FUNCTION_BLOCK basicInversorATV600 (* Inversor ATV600 por Modbus TCP generico: registradores brutos para grandezas e palavras de escrita *)
  (* Standard: 61499-2 *)
  (* Version 1.1, 27/10/2026, Hidryco, Hidryco, 1.1: VELOCIDADE_PCT (leitura) entre LSP 3105 = 0 %% e HSP 3104 = 100 %%. 1.0: Motor_Generico com ATV600 por MODBUSGENTCPS (unit 248): RFR, LCR, UOP, OPR, OTR, LFT e RFRD lidos; LFR e CMD escritos (planilha ATV600 V4.6). *)
  PACKAGE Hidryco.HidrycoLib;
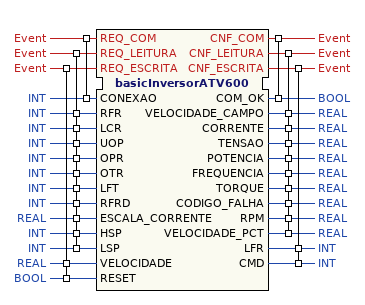
  EVENT_INPUT
    REQ_COM WITH CONEXAO; (* connStatusInt do escravo Modbus *)
    REQ_LEITURA WITH RFR, LCR, UOP, OPR, OTR, LFT, RFRD, ESCALA_CORRENTE, HSP, LSP; (* Nova leitura dos registradores do inversor *)
    REQ_ESCRITA WITH VELOCIDADE, RESET; (* Referencia e reset para o inversor *)
  END_EVENT
  EVENT_OUTPUT
    CNF_COM WITH COM_OK; (* Status de comunicacao *)
    CNF_LEITURA WITH VELOCIDADE_CAMPO, CORRENTE, TENSAO, POTENCIA, FREQUENCIA, TORQUE, CODIGO_FALHA, RPM, VELOCIDADE_PCT; (* Grandezas do inversor *)
    CNF_ESCRITA WITH LFR, CMD; (* Palavras para o inversor *)
  END_EVENT
  VAR_INPUT
    CONEXAO : INT; (* connStatusInt do MODBUSGENTCPS: 1 = online *)
    RFR : INT; (* RFR 3202 - frequencia do motor (0,1 Hz) *)
    LCR : INT; (* LCR 3204 - corrente do motor (UINT, unidade em ESCALA_CORRENTE) *)
    UOP : INT; (* UOP 3208 - tensao do motor (UINT, 1 V) *)
    OPR : INT; (* OPR 3211 - potencia do motor (1 %) *)
    OTR : INT; (* OTR 3205 - torque do motor (0,1 %) *)
    LFT : INT; (* LFT 7121 - ultimo erro ocorrido (WORD) *)
    RFRD : INT; (* RFRD 8604 - velocidade de saida (1 rpm) *)
    ESCALA_CORRENTE : REAL; (* A por unidade do LCR (0,1 = LCR em 0,1 A) *)
    HSP : INT; (* HSP 3104 - velocidade maxima (0,1 Hz) *)
    LSP : INT; (* LSP 3105 - velocidade minima (0,1 Hz) *)
    VELOCIDADE : REAL; (* Referencia de velocidade na unidade de campo (0,1 Hz, cfgSaidaMax = 600) *)
    RESET : BOOL; (* Pulso de reset de falha *)
  END_VAR
  VAR_OUTPUT
    COM_OK : BOOL; (* TRUE = inversor online *)
    VELOCIDADE_CAMPO : REAL; (* Velocidade real na unidade de campo (RFR em 0,1 Hz) *)
    CORRENTE : REAL; (* Corrente (A) *)
    TENSAO : REAL; (* Tensao do motor (V) *)
    POTENCIA : REAL; (* Potencia do motor (%) *)
    FREQUENCIA : REAL; (* Frequencia (Hz) *)
    TORQUE : REAL; (* Torque (%) *)
    CODIGO_FALHA : REAL; (* Ultimo codigo de erro (LFT) *)
    RPM : REAL; (* Rotacao (rpm) *)
    VELOCIDADE_PCT : REAL; (* Velocidade (%) so leitura: 0 % no LSP, 100 % no HSP *)
    LFR : INT; (* LFR 8502 - referencia de frequencia (0,1 Hz) *)
    CMD : INT; (* CMD 8501 - palavra de comando (bit 7 = reset de falha) *)
  END_VAR
  VAR
    r : REAL; (* Auxiliar UINT -> REAL *)
  END_VAR
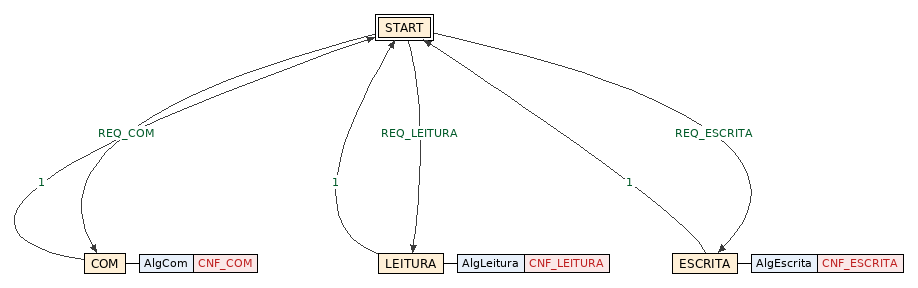
  EC_STATES
    START; (* Initial State *)
    COM : AlgCom -> CNF_COM;
    LEITURA : AlgLeitura -> CNF_LEITURA;
    ESCRITA : AlgEscrita -> CNF_ESCRITA;
  END_STATES
  EC_TRANSITIONS
    START TO COM := REQ_COM;
    COM TO START := 1;
    START TO LEITURA := REQ_LEITURA;
    LEITURA TO START := 1;
    START TO ESCRITA := REQ_ESCRITA;
    ESCRITA TO START := 1;
  END_TRANSITIONS
  ALGORITHM AlgCom IN ST:
(* connStatusInt do escravo Modbus: 1 = online *)
COM_OK := (CONEXAO = 1);
  END_ALGORITHM
  ALGORITHM AlgLeitura IN ST:
(* Registradores do ATV600 (logic addresses da planilha ATV600 V4.6). LCR, UOP e LFT sao UINT/WORD: lidos em INT,
   voltam para 0..65535. A velocidade fica em 0,1 Hz (unidade de campo do Motor_Generico, cfgSaidaMax = 600). *)
VELOCIDADE_CAMPO := INT_TO_REAL(RFR);
FREQUENCIA := INT_TO_REAL(RFR) / 10.0;
r := INT_TO_REAL(LCR);
IF r < 0.0 THEN
    r := r + 65536.0;
END_IF;
CORRENTE := r * ESCALA_CORRENTE;
r := INT_TO_REAL(UOP);
IF r < 0.0 THEN
    r := r + 65536.0;
END_IF;
TENSAO := r;
POTENCIA := INT_TO_REAL(OPR);
TORQUE := INT_TO_REAL(OTR) / 10.0;
r := INT_TO_REAL(LFT);
IF r < 0.0 THEN
    r := r + 65536.0;
END_IF;
CODIGO_FALHA := r;
RPM := INT_TO_REAL(RFRD);
(* Velocidade so para leitura: 0 % no LSP e 100 % no HSP do inversor (parado ou abaixo do LSP = 0 %) *)
IF HSP > LSP THEN
    VELOCIDADE_PCT := LIMIT(0.0, INT_TO_REAL(RFR - LSP) * 100.0 / INT_TO_REAL(HSP - LSP), 100.0);
ELSE
    VELOCIDADE_PCT := 0.0;
END_IF;
  END_ALGORITHM
  ALGORITHM AlgEscrita IN ST:
(* LFR em 0,1 Hz (faixa da planilha -5000..5000); CMD bit 7 = reset de falha, 0 fora do pulso.
   A partida do motor continua pela saida digital (cmdAcionamento). *)
LFR := REAL_TO_INT(LIMIT(-5000.0, VELOCIDADE, 5000.0));
IF RESET THEN
    CMD := 128;
ELSE
    CMD := 0;
END_IF;
  END_ALGORITHM
END_FUNCTION_BLOCK
